Staubli VAL3: getProgList.pgx

public program getProgList(string& x_sList[])
  local string l_sKey
begin
  resize(x_sList,1,1)
  l_sKey=first(progTemp:pProgItem)

  while l_sKey!=""
    x_sList[size(x_sList)-1]=l_sKey
    insert(x_sList[size(x_sList)])
    l_sKey=next(progTemp:pProgItem[l_sKey])
  endWhile
end
